(* IEC 61131-3 sources: llm-plc-st-eval/data/definitivo/qwen2.5-coder_14b/A1/few_shot, 3 files *)

(* ---- ejec_1.st ---- *)
FUNCTION_BLOCK FB_PID
VAR_INPUT
    SP : REAL; (* Consigna *)
    PV : REAL; (* Variable de proceso *)
    Kp : REAL; (* Ganancia proporcional *)
    Ti : REAL; (* Tiempo integral en segundos *)
    Td : REAL; (* Tiempo derivativo en segundos *)
    ciclo : TIME; (* Ciclo de muestreo *)
END_VAR
VAR_OUTPUT
    CV : REAL; (* Salida del controlador PID *)
END_VAR
VAR
    e : REAL; (* Error *)
    e_prev : REAL; (* Error previo *)
    integral : REAL; (* Integral del error *)
    derivativa : REAL; (* Derivada del error *)
    dt : TIME; (* Intervalo de tiempo entre ejecuciones *)
END_VAR

(* Calculo del error *)
e := SP - PV;

(* Calculo de la derivativa *)
dt := ciclo;
derivativa := (e - e_prev) / REAL_TO_TIME(dt);

(* Calculo de la integral *)
IF Ti > 0.0 THEN
    integral := integral + (e * REAL_TO_TIME(dt)) / Ti;
ELSE
    integral := 0.0; (* Desactiva la acción integral *)
END_IF;

(* Anti-windup por clamping *)
IF CV >= 100.0 THEN
    IF e > 0.0 THEN
        integral := integral - e * REAL_TO_TIME(dt) / Ti; (* No acumula error positivo *)
    END_IF;
ELSIF CV <= 0.0 THEN
    IF e < 0.0 THEN
        integral := integral - e * REAL_TO_TIME(dt) / Ti; (* No acumula error negativo *)
    END_IF;
END_IF;

(* Calculo de la salida CV *)
CV := Kp * (e + integral + Td * derivativa);

(* Limita la salida CV al rango 0.0 a 100.0 *)
IF CV > 100.0 THEN
    CV := 100.0;
ELSIF CV < 0.0 THEN
    CV := 0.0;
END_IF;

(* Actualiza el error previo *)
e_prev := e;
END_FUNCTION_BLOCK

(* ---- ejec_2.st ---- *)
FUNCTION_BLOCK FB_PID
VAR_INPUT
    SP : REAL; (* Setpoint *)
    PV : REAL; (* Process Variable *)
    Kp : REAL; (* Proportional Gain *)
    Ti : REAL; (* Integral Time in seconds *)
    Td : REAL; (* Derivative Time in seconds *)
    ciclo : TIME; (* Sampling Cycle *)
END_VAR
VAR_OUTPUT
    CV : REAL; (* Control Variable, 0.0 to 100.0 *)
END_VAR
VAR
    e : REAL; (* Error *)
    ePrev : REAL; (* Previous Error *)
    integral : REAL; (* Integral of Error *)
    derivativa : REAL; (* Derivative of Error *)
    dt : TIME; (* Time Difference *)
END_VAR

(* Calculate the error *)
e := SP - PV;

(* Calculate the derivative of the error *)
dt := ciclo;
derivativa := (e - ePrev) / REAL_TO_TIME(dt);

(* Calculate the integral of the error *)
IF Ti > 0.0 THEN
    integral := integral + (e * REAL_TO_TIME(ciclo)) / Ti;
ELSE
    integral := 0.0; (* Integral action disabled *)
END_IF;

(* Anti-windup by clamping *)
IF CV >= 100.0 THEN
    IF e > 0.0 THEN
        integral := integral - e * REAL_TO_TIME(ciclo) / Ti; (* Prevent integral windup *)
    END_IF;
ELSIF CV <= 0.0 THEN
    IF e < 0.0 THEN
        integral := integral - e * REAL_TO_TIME(ciclo) / Ti; (* Prevent integral windup *)
    END_IF;
END_IF;

(* Calculate the control variable *)
CV := Kp * (e + integral + Td * derivativa);

(* Clamp the control variable to the range 0.0 to 100.0 *)
IF CV > 100.0 THEN
    CV := 100.0;
ELSIF CV < 0.0 THEN
    CV := 0.0;
END_IF;

(* Update previous error *)
ePrev := e;
END_FUNCTION_BLOCK

(* ---- ejec_3.st ---- *)
FUNCTION_BLOCK FB_PID
VAR_INPUT
    SP : REAL; (* Consigna *)
    PV : REAL; (* Variable de proceso *)
    Kp : REAL; (* Ganancia proporcional *)
    Ti : REAL; (* Tiempo integral en segundos *)
    Td : REAL; (* Tiempo derivativo en segundos *)
    ciclo : TIME; (* Ciclo de muestreo *)
END_VAR
VAR_OUTPUT
    CV : REAL; (* Salida del controlador PID, porcentaje de mando *)
END_VAR
VAR
    e : REAL; (* Error *)
    e_prev : REAL; (* Error anterior *)
    integral : REAL; (* Integral del error *)
    derivada : REAL; (* Derivada del error *)
    dt : TIME; (* Intervalo de tiempo entre ejecuciones *)
END_VAR

(* Calculo del error *)
e := SP - PV;

(* Calculo de la derivada *)
dt := ciclo;
derivada := (e - e_prev) / REAL_TO_TIME(dt);

(* Calculo de la integral *)
IF Ti > 0.0 THEN
    integral := integral + (e * REAL_TO_TIME(dt)) / Ti;
ELSE
    integral := 0.0; (* Desactiva la acción integral *)
END_IF;

(* Anti-windup por clamping *)
IF CV >= 100.0 THEN
    IF e > 0.0 THEN
        integral := integral - (e * REAL_TO_TIME(dt)) / Ti; (* No acumula error positivo *)
    END_IF;
ELSIF CV <= 0.0 THEN
    IF e < 0.0 THEN
        integral := integral - (e * REAL_TO_TIME(dt)) / Ti; (* No acumula error negativo *)
    END_IF;
END_IF;

(* Calculo de la salida CV *)
CV := Kp * (e + integral + Td * derivada);

(* Limita CV al rango 0.0 a 100.0 *)
IF CV > 100.0 THEN
    CV := 100.0;
ELSIF CV < 0.0 THEN
    CV := 0.0;
END_IF;

(* Actualiza el error anterior *)
e_prev := e;
END_FUNCTION_BLOCK
